Fanuc KAREL source: kb00198.KL

-- PROVISIONAL review KL for V1013-1; original PC SHA256 b160ff4c530e0839d2e52cb6dbf1ea310eac31607527ec72f6c719e7ea2fcdb7
-- Incomplete behavior may be omitted. Consult companion uncertainty JSON. Do not deploy.
PROGRAM KB00198
%NOLOCKGROUP
BEGIN
  -- UNRESOLVED_PC offsets 5-14; opcodes 3F,75
  -- UNRESOLVED_PC offsets 19-26; opcodes 9D,23
  -- UNRESOLVED_PC offsets 31-38; opcodes 9D,23
  -- UNRESOLVED_PC offsets 43-79; opcodes 27,22,22,2A,22,22,22,31
  -- UNRESOLVED_PC offsets 84-88; opcodes 7F
END KB00198
